(* IEC 61131-3 sources: Test-Git_ESME26/TestProgettoESME_26.fbsproj/TemplateFullProgrammingFramework_Migration.device.xml.v3^/Plc Logic.plclogic.xml.v3^/Application.application.xml.v3^/Sercos_Template/WriteIDN/FB_Set230VModeAsync.fb.st^, 2 files *)

(* ---- Set230VMode.meth.st ---- *)
METHOD Set230VMode : dint
VAR_INPUT
	i_ifSercosIdentificationAccess : SDI.IF_SercosIdentificationAccess;
END_VAR
VAR_OUTPUT
	//q_diResult : DINT;
	q_sDiagMsg : STRING[255];
END_VAR
VAR
	diResult : DINT;
	ifLxm62PowerSupplyAccess : LXM62SI.IF_Lxm62PowerSupplyAccess;
END_VAR

// Check if we have a Lexium62 PowerSupply
IF __QUERYINTERFACE(i_ifSercosIdentificationAccess, ifLxm62PowerSupplyAccess) THEN
	// Set 'PhaseCheckMode' (P-0-0638) to 1 phase (1)
	diResult := FC_SercosWriteIDN(
		i_uiTopoAddr := i_ifSercosIdentificationAccess.SercosIdentification.ConfiguredTopologyAddress,
		i_etSercosParameterType := ET_SercosParameterType.P_Parameter,
		i_uiIDN := 638,
		i_etWriteIDNType := ET_SercosWriteIDNType.WriteUserData,
		i_dwValue := 1);

	IF diResult <> 0 THEN
		q_sDiagMsg := 'Set $'PhaseCheckMode$' to $'230 V / 1$' on PowerSupply failed.';
		Set230VMode := diResult;
		RETURN;
	END_IF
END_IF

// Set 'MainsVoltageMode' (P-0-1021) to 230V (1) - for PowerSupply and Drives
diResult := FC_SercosWriteIDN(
	i_uiTopoAddr := i_ifSercosIdentificationAccess.SercosIdentification.ConfiguredTopologyAddress,
	i_etSercosParameterType := ET_SercosParameterType.P_Parameter,
	i_uiIDN := 1021,
	i_etWriteIDNType := ET_SercosWriteIDNType.WriteUserData,
	i_dwValue := 1);

IF diResult <> 0 THEN
	q_sDiagMsg := 'Set $'MainsVoltageMode$' to $'230 V / 1$' on Sercos device failed.';
	Set230VMode := diResult;
	RETURN;
END_IF

(* ---- xDone.prop.st ---- *)
PROPERTY xDone : BOOL
__GETTERDECLARATION__
VAR
END_VAR
__GETTERIMPLEMENTATION__
xDone := xDone_loc;
__SETTERDECLARATION__
VAR
END_VAR
__SETTERIMPLEMENTATION__
xDone_loc := xDone;
